(* IEC 61131-3 sources: kns-port-domestic/targets/astra/src/POUs/Station/FB_Annunciator, 2 files *)

(* ---- FB_Annunciator.decl.st ---- *)
// Назначение: местная сигнализация (04 §14): сирена HA1 — новая неквитированная тревога High или
//             Critical, выключается кнопкой HS502, командой «Звук» или квитированием, новая
//             тревога включает снова; лампа HL1 — мигает 1 Гц при неквитированных Medium и выше,
//             горит при активных квитированных; реле K1 «Общая авария» — под напряжением в норме,
//             обесточено при активной High или Critical (принцип «отказ — сигнал»).
// Автор:      kr0nsch
// Версия:     0.1.0
// Документ:   docs/DESIGN.md, раздел 6.12; docs/04_algorithms.md, раздел 14
FUNCTION_BLOCK FB_Annunciator
VAR_INPUT
    auiUnack      : ARRAY[1..GVL_Const.ALM_PRIO_COUNT] OF UINT;   // Low…Critical (FB_AlarmSummary)
    auiActive     : ARRAY[1..GVL_Const.ALM_PRIO_COUNT] OF UINT;
    udiNewHighSeq : UDINT;          // растёт на каждую новую неквитированную High/Critical
    xSilence      : BOOL;           // импульс: фронт HS502 OR stStationCmd.xSilence
    itfTime       : PL.I_TimeSource;
END_VAR
VAR_OUTPUT
    xHorn        : BOOL;            // → GVL_IO.xHA1
    xLamp        : BOOL;            // → GVL_IO.xHL1: мигает 1 Гц при неквитированных Medium+, горит при активных
    xK1Energized : BOOL;            // → GVL_IO.xK1: TRUE — норма, FALSE — активна High/Critical
END_VAR
VAR
    udiSeqPrev   : UDINT;           // udiNewHighSeq прошлого вызова
    xFirstCall   : BOOL := TRUE;    // первый вызов: счётчик сводки принимается как есть
    xBlinking    : BOOL;            // лампа в режиме мигания (прошлый вызов)
    ltBlinkStart : LTIME;           // начало мигания: фаза «горит»
    fbSysTime    : PL.FB_SystemTime;    // запасной источник времени (itfTime = 0)
END_VAR
VAR_TEMP
    uiPrio      : UINT;             // индекс приоритета
    uiUnackMed  : UINT;             // неквитированных Medium и выше
    uiUnackHigh : UINT;             // неквитированных High и выше
    uiActMed    : UINT;             // активных Medium и выше
    uiActHigh   : UINT;             // активных High и выше
    ltNow       : LTIME;            // время этого вызова
    uliHalf     : ULINT;            // полупериод мигания, нс
END_VAR

(* ---- FB_Annunciator.impl.st ---- *)
// 1. Счётчики по приоритетам (индекс — значение E_AlarmPriority: Low = 1 … Critical = 4)
uiUnackMed := 0;
uiUnackHigh := 0;
uiActMed := 0;
uiActHigh := 0;
FOR uiPrio := TO_UINT(PL.E_AlarmPriority.Medium) TO GVL_Const.ALM_PRIO_COUNT DO
    uiUnackMed := uiUnackMed + auiUnack[uiPrio];
    uiActMed := uiActMed + auiActive[uiPrio];
    IF uiPrio >= TO_UINT(PL.E_AlarmPriority.High) THEN
        uiUnackHigh := uiUnackHigh + auiUnack[uiPrio];
        uiActHigh := uiActHigh + auiActive[uiPrio];
    END_IF
END_FOR

// 2. Сирена: «Звук» выключает, новая High/Critical включает снова (новая старше команды того же
//    цикла), квитирование всех High/Critical — выключает
IF xFirstCall THEN
    udiSeqPrev := udiNewHighSeq;
END_IF
IF xSilence THEN
    xHorn := FALSE;
END_IF
IF udiNewHighSeq <> udiSeqPrev THEN
    xHorn := TRUE;
END_IF
IF uiUnackHigh = 0 THEN
    xHorn := FALSE;
END_IF
udiSeqPrev := udiNewHighSeq;

// 3. Лампа: мигание 1 Гц по времени источника (фаза «горит» — с начала мигания), иначе горит при
//    активных; «время назад» начинает мигание заново
IF itfTime <> 0 THEN
    ltNow := itfTime.Now();
ELSE
    ltNow := fbSysTime.Now();
END_IF
IF uiUnackMed > 0 THEN
    IF NOT xBlinking OR ltNow < ltBlinkStart THEN
        ltBlinkStart := ltNow;
    END_IF
    xBlinking := TRUE;
    // PORT: [types] проверить в Astra.IDE — литералы и преобразования LTIME (C11)
    uliHalf := LTIME_TO_ULINT(TIME_TO_LTIME(GVL_Const.STN_LAMP_HALF_PERIOD));
    IF uliHalf > 0 THEN
        // PORT: [types] проверить в Astra.IDE — литералы и преобразования LTIME (C11)
        xLamp := ((LTIME_TO_ULINT(ltNow - ltBlinkStart) / uliHalf) MOD 2) = 0;
    ELSE
        xLamp := TRUE;
    END_IF
ELSE
    xBlinking := FALSE;
    xLamp := uiActMed > 0;
END_IF

// 4. Реле «Общая авария»: под напряжением в норме
xK1Energized := uiActHigh = 0;
xFirstCall := FALSE;
